// TIA Portal V21 export
ORGANIZATION_BLOCK "PipCyclic"   // OB30, SCL, CyclicInterrupt
{ S7_Optimized_Access := 'TRUE' }
// stored: AutoNumber false
   VAR_INPUT
      Initial_Call : Bool;
      Event_Count : Int;
   END_VAR
BEGIN
   "PipDb".Ob30Count := "PipDb".Ob30Count + 1;
END_ORGANIZATION_BLOCK
